(* IEC 61131-3 sources: rusty/tests/lit/single/builtin, 8 files *)

(* ---- abs_unsigned.st ---- *)
// RUN: (%COMPILE %s && %RUN) | %CHECK %s
//
// ABS with an unsigned argument binds to the ABS__U* builtins and returns the
// value unchanged instead of calling a non-existent library monomorph
// (previously a crash at runtime). Signed and float arguments still call the
// library implementations.

FUNCTION main
VAR
    s   : SINT  := SINT#-128;
    i   : INT   := INT#-3;
    d   : DINT  := DINT#-10;
    l   : LINT  := LINT#-1234567890123;
    u8  : USINT := USINT#200;
    u16 : UINT  := UINT#5;
    u32 : UDINT := UDINT#4000000000;
    u64 : ULINT := ULINT#42;
    r   : REAL  := REAL#-2.0;
    lr  : LREAL := LREAL#-9.5;
END_VAR

// ABS(INT_MIN) wraps to INT_MIN
// CHECK: s=-128
printf('s=%d$N', ABS(s));

// CHECK: i=3
printf('i=%d$N', ABS(i));

// CHECK: d=10
printf('d=%d$N', ABS(d));

// CHECK: l=1234567890123
printf('l=%lld$N', ABS(l));

// CHECK: u8=200
printf('u8=%d$N', ABS(u8));

// CHECK: u16=5
printf('u16=%d$N', ABS(u16));

// CHECK: u32=4000000000
printf('u32=%u$N', ABS(u32));

// CHECK: u64=42
printf('u64=%llu$N', ABS(u64));

// CHECK: r=2.0
printf('r=%.1f$N', ABS(r));

// CHECK: lr=9.5
printf('lr=%.1f$N', ABS(lr));

// explicit calls to the library monomorphs still link against the stdlib
// CHECK: lib=7
printf('lib=%d$N', ABS__DINT(DINT#-7));
END_FUNCTION

(* ---- abs_unsigned_warning.st ---- *)
// RUN: %COMPILE %s 2>&1 | %CHECK %s
//
// ABS of an unsigned value has no effect and reports a warning for each call.

FUNCTION main
VAR
    u8  : USINT;
    u16 : UINT;
    u32 : UDINT;
    u64 : ULINT;
    res : ULINT;
END_VAR

// CHECK: {{.*}}warning[E150]{{.*}}ABS on a value of unsigned type 'USINT' has no effect{{.*}}
res := ABS(u8);

// CHECK: {{.*}}warning[E150]{{.*}}ABS on a value of unsigned type 'UINT' has no effect{{.*}}
res := ABS(u16);

// CHECK: {{.*}}warning[E150]{{.*}}ABS on a value of unsigned type 'UDINT' has no effect{{.*}}
res := ABS(u32);

// CHECK: {{.*}}warning[E150]{{.*}}ABS on a value of unsigned type 'ULINT' has no effect{{.*}}
res := ABS(u64);
END_FUNCTION

(* ---- adr_ptr_arith_runtime.st ---- *)
// RUN: (%COMPILE %s && %RUN) | %CHECK %s
//
// `ADR(x) + N` is byte-stride pointer arithmetic — `ADR` is declared to
// return LWORD, so the `+` flows through the integer-arithmetic path; the
// receiver pointer ends up `N` bytes past the operand. Regression for #1749
// (previously panicked in `create_llvm_int_binary_expression`).

FUNCTION main
VAR
    arr : ARRAY[0..7] OF BYTE := [0, 0, 0, 0, 0, 0, 0, 0];
    pt  : REF_TO BYTE;
END_VAR

pt := ADR(arr) + 4;
pt^ := BYTE#16#AB;

// CHECK: arr[4]=171
printf('arr[4]=%d$N', arr[4]);

pt := ADR(arr) + 7;
pt^ := BYTE#16#5C;

// CHECK: arr[7]=92
printf('arr[7]=%d$N', arr[7]);

// Subtraction flows through the same path: take a pointer past the end
// and walk back. Writing to arr[2] via `ADR(arr[6]) - 4`.
pt := ADR(arr[6]) - 4;
pt^ := BYTE#16#11;

// CHECK: arr[2]=17
printf('arr[2]=%d$N', arr[2]);
END_FUNCTION

(* ---- datetime_arithmetic_operators.st ---- *)
// RUN: (%COMPILE %s && %RUN) | %CHECK %s
// The operators on date and time operands: a time of day wraps at midnight, a real factor is
// applied as such, and every other combination is the plain nanosecond arithmetic

FUNCTION main
    VAR
        t1, t2, t : TIME;
        tod : TOD;
        d1, d2 : DATE;
        dt1, dt2 : DT;
        ltod : LTOD;
        lt : LTIME;
    END_VAR
    t1 := T#1s; t2 := T#500ms; t := t1 + t2;
    printf('%s$N', REF(TIME_TO_STRING(t)));                                         // CHECK: T#1s500ms
    tod := TOD#23:59:50 + T#20s;
    printf('%s %lld$N', REF(TOD_TO_STRING(tod)), tod);                              // CHECK: TOD#00:00:10 10000000000
    tod := TOD#00:00:10 - T#20s;
    printf('%s %lld$N', REF(TOD_TO_STRING(tod)), tod);                              // CHECK: TOD#23:59:50 86390000000000
    dt1 := DT#2024-01-15-12:30:00 + T#5s;
    printf('%s$N', REF(DT_TO_STRING(dt1)));                                         // CHECK: DT#2024-01-15-12:30:05
    t1 := T#10s; t2 := T#3s; t := t1 - t2;
    printf('%s$N', REF(TIME_TO_STRING(t)));                                         // CHECK: T#7s
    d1 := D#2024-01-15; d2 := D#2024-01-10; t := d1 - d2;
    printf('%s$N', REF(TIME_TO_STRING(t)));                                         // CHECK: T#5d
    t := TOD#10:30:00 - TOD#10:20:00;
    printf('%s$N', REF(TIME_TO_STRING(t)));                                         // CHECK: T#10m
    dt1 := DT#2024-01-15-12:30:10; dt2 := DT#2024-01-15-12:30:00; t := dt1 - dt2;
    printf('%s$N', REF(TIME_TO_STRING(t)));                                         // CHECK: T#10s
    t := t1 * 3;
    printf('%s$N', REF(TIME_TO_STRING(t)));                                         // CHECK: T#30s
    t := 2 * t1;
    printf('%s$N', REF(TIME_TO_STRING(t)));                                         // CHECK: T#20s
    t := t1 / 4;
    printf('%s$N', REF(TIME_TO_STRING(t)));                                         // CHECK: T#2s500ms
    t := t1 * 1.5;
    printf('%s$N', REF(TIME_TO_STRING(t)));                                         // CHECK: T#15s
    t := 1.5 * t1;
    printf('%s$N', REF(TIME_TO_STRING(t)));                                         // CHECK: T#15s
    t := t1 / 2.5;
    printf('%s$N', REF(TIME_TO_STRING(t)));                                         // CHECK: T#4s
    ltod := LTOD#23:59:50 + LTIME#20s;
    printf('%s %lld$N', REF(LTOD_TO_STRING(ltod)), ltod);                           // CHECK: LTOD#00:00:10 10000000000
    lt := LTIME#10s * 1.5;
    printf('%s$N', REF(LTIME_TO_STRING(lt)));                                       // CHECK: LTIME#15s
    t := t1 + 5;
    printf('%s$N', REF(TIME_TO_STRING(t)));                                         // CHECK: T#10s5ns
    dt1 := DT#2027-05-05-22:30:15 + T#20s + T#20s + T#2h555s;
    printf('%s$N', REF(DT_TO_STRING(dt1)));                                         // CHECK: DT#2027-05-06-00:40:10
END_FUNCTION

(* ---- shl_and_shr_must_cast_left_and_right_correctly.st ---- *)
// RUN: (%COMPILE %s && %RUN) | %CHECK %s

// SHL and SHR must cast left and right correctly
FUNCTION main
VAR
    value : BYTE;
END_VAR

value := BIT_LOAD_B2(BYTE#255, TRUE, 2, 2);

// CHECK: 255
printf('%d$N', value);

value := BIT_LOAD_B2(BYTE#255, FALSE, 2, 2);

// CHECK: 243
printf('%d$N', value);

END_FUNCTION

FUNCTION BIT_LOAD_B2 : BYTE
VAR_INPUT
	I : BYTE;
	D : BOOL;
	P : INT;
	N : INT;
END_VAR
VAR
    result : BYTE;
END_VAR

IF D THEN
	BIT_LOAD_B2 := ROL(SHR(BYTE#255, 8 - N) OR ROR(I, P), P);
ELSE
	BIT_LOAD_B2 := ROL(SHL(BYTE#255, N) AND ROR(I, P), P);
END_IF;

END_FUNCTION

(* ---- shl_must_be_usable_with_integers.st ---- *)
// RUN: (%COMPILE %s && %RUN) | %CHECK %s

// SHL must be usable with integers
FUNCTION main
VAR
    a : INT;
END_VAR
a := SHL(21,2);

// CHECK: 84
printf('%d$N', a);
END_FUNCTION

(* ---- shr_must_be_usable_with_integers.st ---- *)
// RUN: (%COMPILE %s && %RUN) | %CHECK %s

// SHR must be usable with integers
FUNCTION main
VAR
    a : INT;
END_VAR
a := SHR(21,2);

// CHECK: 5
printf('%d$N', a);
END_FUNCTION

(* ---- shr_unsigned_byte_logical_shift.st ---- *)
// RUN: (%COMPILE %s && %RUN) | %CHECK %s

// SHR on unsigned BYTE must use logical shift (zero-fill), not arithmetic shift
FUNCTION main
VAR
    b : BYTE;
    s : SINT;
END_VAR
b := SHR(BYTE#251, SINT#1);

// CHECK: 125
printf('%d$N', b);

s := SHR(SINT#-4, SINT#1);

// CHECK: -2
printf('%d$N', s);
END_FUNCTION
